// TIA Portal V20 export
// export: Created 2026-10-12T16:46:21.4347175Z, ExportSetting WithDefaults, DisplayName Totally Integrated Automation Portal, DisplayVersion V20 Update 6, DisplayName TIA Portal Openness, DisplayVersion V20 Update 6, DisplayName TIA Portal Version Control Interface, DisplayVersion V20 Update 6, DisplayName SINAMICS Startdrive Advanced, DisplayVersion V20 SP1 Update 2, DisplayName SINAMICS Startdrive G110M, G120, G120C, G120D, G120P, G115D, DisplayVersion V20 SP1 Update 2, DisplayName SINAMICS Startdrive G130, G150, S120, S150, SINAMICS MV, G220, S200, S210, DisplayVersion V20 SP1 Update 2, DisplayName STEP 7 Professional, DisplayVersion V20 Update 6, DisplayName STEP 7 Safety, DisplayVersion V20 Update 2, DisplayName WinCC Basic/Comfort/Advanced, DisplayVersion V20 Update 6, DisplayName WinCC Professional, DisplayVersion V20 Update 6, DisplayName WinCC Unified, DisplayVersion V20 Update 6
DATA_BLOCK "FB_Bad_DB"   // DB41
VERSION : 0.2
// stored: AutoNumber true, DBAccessibleFromOPCUA true, DBAccessibleFromWebserver true, InstanceOfName FB_Bad, InstanceOfType FB
"FB_Bad"
   // VAR_INPUT
   //    Blink_Takt : Bool;
   //    Lampentest : Bool;
   //    Blink_Zaehler : Int;
   //    Not_Halt_Aktiv : Bool;
   //    Zustand : Int;
   //    BadNr : Int;
   // END_VAR
   // VAR_IN_OUT
   //    Bad_Konfig : "UDT_Bad_Konfig";
   //    Auftraege : Array[0..9] of "UDT_Prozessroute";
   //    Handbetrieb : "UDT_Handbetrieb";
   //    Leerlauf : "UDT_Peripherie_Soll";
   //    Standby : "UDT_Peripherie_Soll";
   // END_VAR
   // VAR
   //    Timer_WT { S7_SetPoint := 'True'} : Array[1..3] of TON_TIME;
   //    Timer_FU_Pause { S7_SetPoint := 'True'} : TON_TIME;
   //    Timer_FU_Pumpe_Stoerung { S7_SetPoint := 'True'} : TON_TIME;
   //    Timer_FU_WB1_Stoerung { S7_SetPoint := 'True'} : TON_TIME;
   //    Timer_FU_WB2_Stoerung { S7_SetPoint := 'True'} : TON_TIME;
   //    M_Ein_Any_Alt : Bool;
   //    M_Ent_Any_Alt : Bool;
   // END_VAR
BEGIN
END_DATA_BLOCK
